RoboDK station: kuka_frame.rdk

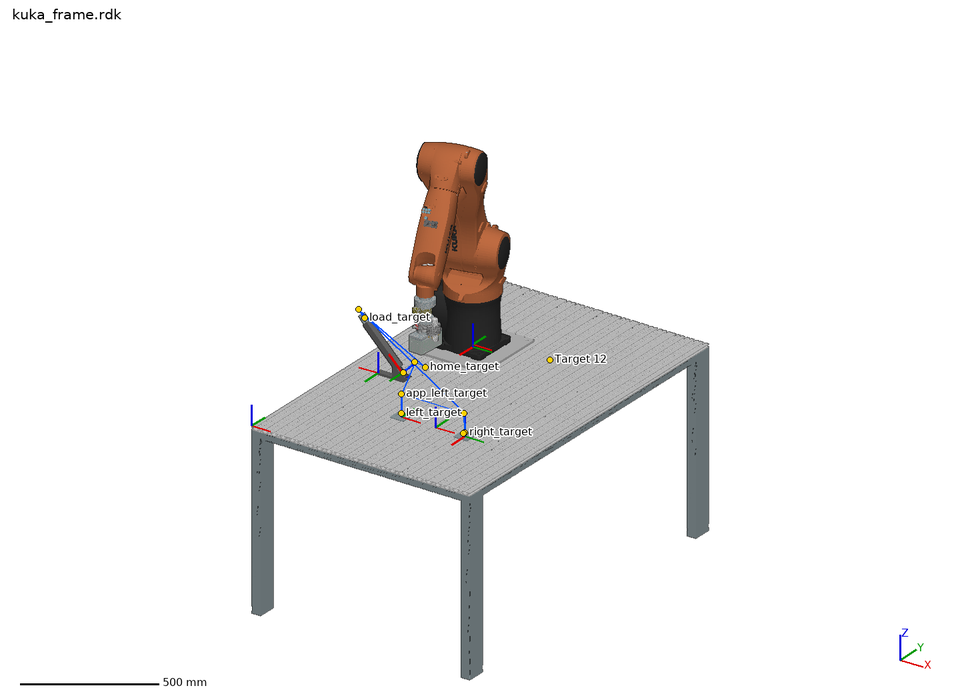
[picture v0: the station drawn from its stored meshes, robots at their saved joint values, targets as dots, program paths as lines]
Station kuka_frame(vansh2) (saved by RoboDK 5.8.0). Poses are relative to the parent item; angles as X-Y-Z fixed-axis rotations.
Station parameters (name, value as stored): LIN64
  - frame table_frame at (0, 0, 0) mm
    - object table_object at (0, 0, 0) mm, size 960.1 x 1500 x 750 mm, geometry from table_object.sld
    - frame base_plate_frame at (280, 990, 0) mm, rotated rx 0 ry 0 rz -90 deg
      - object base_plate_object at (0, 0, 0) mm, size 320 x 320 x 10 mm, geometry from base_plate_object.sld
    - frame slider_frame at (125, 617, 0) mm, rotated rx 0 ry 0 rz 180 deg
      - object slider_object at (0, 0, 0) mm, size 198.7 x 26 x 198.7 mm, 1 curves, geometry from slider_object.sld
    - frame slider_parts_frame at (232.7, 617, 30.7) mm, rotated rx 0 ry -45 rz 180 deg
    - frame pickanddrop at (550, 370, 0) mm
    - frame right_frame at (680, 370, 0) mm, rotated rx 0 ry 0 rz -90 deg
      - object right_plate_object at (0, 0, 0) mm, size 60 x 60 x 9 mm, 1 curves, geometry from right_plate_object.sld
    - frame left_frame at (400, 370, 0) mm
      - object left_plate_object at (0, 0, 0) mm, size 60 x 60 x 9 mm, 1 curves, geometry from left_plate_object.sld
    - frame kuka_frame at (280, 990, 10) mm
      - robot KUKA KR 6 R900 sixx: 6 axes, payload 6 kg, reach 901 mm, repeatability 0.03 mm, weight 52 kg
          modified DH rows (alpha deg, a mm, theta deg, d mm): 0, 0, 0, 400; -90, 25, 0, 0; 0, 455, -90, 0; -90, 35, 0, 420; 90, 0, 0, 0; -90, 0, 180, 80
          joint limits [-170, -190, -120, -185, -120, -350] to [170, 45, 156, 185, 120, 350]; home [0, -90, 90, 0, 0, 0]; saved at [75.683, -66.176, 119.978, 0, 36.199, -61.317]
        - robot gripper: 1 axes
            joint limits [0] to [50]; home [0]; saved at [50]
        - tool gripper_tcp, TCP at (0, 0, 288) mm, rotated rx 0 ry 0 rz 43 deg
    - target home_target (Cartesian target) at (399.96, 519.99, 139.97) mm, rotated rx -180 ry 0 rz 0 deg; joints [75.683, -66.176, 119.978, 0, 36.199, -61.317] of KUKA KR 6 R900 sixx
    - target left_target (Cartesian target) at (400, 370, 15) mm, rotated rx -180 ry 0 rz 0 deg; joints [79.046, -41.366, 97.165, 0, 34.201, -57.954] of KUKA KR 6 R900 sixx
    - target app_left_target (Cartesian target) at (400, 370, 93) mm, rotated rx -180 ry 0 rz 0 deg; joints [79.046, -48.593, 96.885, 0, 41.708, -57.954] of KUKA KR 6 R900 sixx
    - target right_target (Cartesian target) at (680, 370, 15) mm, rotated rx -180 ry 0 rz -90 deg; joints [57.171, -31.816, 75.866, 0, 45.949, -169.829] of KUKA KR 6 R900 sixx
    - target app_right_target (Cartesian target) at (676.53, 370, 93) mm, rotated rx -180 ry 0 rz -180 deg; joints [57.398, -38.147, 75.992, 0, 52.155, 100.398] of KUKA KR 6 R900 sixx
    - target slider_part_target (Cartesian target) at (234.82, 617, 32.82) mm, rotated rx 180 ry 45 rz 0 deg; joints [60.036, -41.203, 127.341, 56.857, 47.023, -132.424] of KUKA KR 6 R900 sixx
    - target app_sliderpart_target (Cartesian target) at (286, 617, 88.78) mm, rotated rx -180 ry 50 rz 0 deg; joints [52.337, -44.49, 122.484, 45.711, 57.903, -125.791] of KUKA KR 6 R900 sixx
    - target load_target (Cartesian target) at (66.24, 617, 203.91) mm, rotated rx -180 ry 50 rz 0 deg; joints [79.647, -66.13, 137.097, 65.731, 55.754, -114.165] of KUKA KR 6 R900 sixx
    - target app_load_target (Cartesian target) at (38.79, 617, 231.21) mm, rotated rx 180 ry 49 rz 0 deg; joints [84.408, -71.376, 137.116, 65.861, 55.395, -107.211] of KUKA KR 6 R900 sixx
    - target open_grip (joint target) at (399.96, 519.99, -148.03) mm, rotated rx -180 ry 0 rz -43 deg; joints [50] of gripper
    - target close_grippertarget (joint target) at (399.96, 519.99, -148.03) mm, rotated rx -180 ry 0 rz -43 deg; joints [20, -66.176, 119.978, -180, -36.199, 118.683] of gripper
    - target Target 12 (Cartesian target) at (735.82, 824.09, 139.97) mm, rotated rx -180 ry 0 rz 55.68 deg; joints [20, -66.176, 119.978, 0, 36.199, 298.683] of KUKA KR 6 R900 sixx
    - target Target 13 (Cartesian target) at (735.82, 824.09, 139.97) mm, rotated rx -180 ry 0 rz 55.68 deg; joints [20, -66.176, 119.978, 0, 36.199, 298.683] of KUKA KR 6 R900 sixx
    - target Target 14 (Cartesian target) at (735.82, 824.09, 139.97) mm, rotated rx -180 ry 0 rz 55.68 deg; joints [20, -66.176, 119.978, 0, 36.199, 298.683] of KUKA KR 6 R900 sixx
    - target Target 15 (Cartesian target) at (735.82, 824.09, 139.97) mm, rotated rx -180 ry 0 rz 55.68 deg; joints [20, -66.176, 119.978, 0, 36.199, 298.683] of KUKA KR 6 R900 sixx
    - target Target 16 (Cartesian target) at (735.82, 824.09, 139.97) mm, rotated rx -180 ry 0 rz 55.68 deg; joints [20, -66.176, 119.978, 0, 36.199, 298.683] of KUKA KR 6 R900 sixx
    - target Target 17 (Cartesian target) at (735.82, 824.09, 139.97) mm, rotated rx -180 ry 0 rz 55.68 deg; joints [20, -66.176, 119.978, 0, 36.199, 298.683] of KUKA KR 6 R900 sixx
    - target Target 18 (Cartesian target) at (735.82, 824.09, 139.97) mm, rotated rx -180 ry 0 rz 55.68 deg; joints [20, -66.176, 119.978, 0, 36.199, 298.683] of KUKA KR 6 R900 sixx
    - target Target 19 (Cartesian target) at (735.82, 824.09, 139.97) mm, rotated rx -180 ry 0 rz 55.68 deg; joints [20, -66.176, 119.978, 0, 36.199, 298.683] of KUKA KR 6 R900 sixx
    - target Target 20 (Cartesian target) at (735.82, 824.09, 139.97) mm, rotated rx -180 ry 0 rz 55.68 deg; joints [20, -66.176, 119.978, 0, 36.199, 298.683] of KUKA KR 6 R900 sixx
    - target Target 21 (Cartesian target) at (735.82, 824.09, 139.97) mm, rotated rx -180 ry 0 rz 55.68 deg; joints [20, -66.176, 119.978, 0, 36.199, 298.683] of KUKA KR 6 R900 sixx
    - target Target 22 (Cartesian target) at (735.82, 824.09, 139.97) mm, rotated rx -180 ry 0 rz 55.68 deg; joints [20, -66.176, 119.978, 0, 36.199, 298.683] of KUKA KR 6 R900 sixx
    - target Target 23 (Cartesian target) at (735.82, 824.09, 139.97) mm, rotated rx -180 ry 0 rz 55.68 deg; joints [20, -66.176, 119.978, 0, 36.199, 298.683] of KUKA KR 6 R900 sixx
    - target Target 24 (Cartesian target) at (735.82, 824.09, 139.97) mm, rotated rx -180 ry 0 rz 55.68 deg; joints [20, -66.176, 119.978, 0, 36.199, 298.683] of KUKA KR 6 R900 sixx
    - target Target 25 (Cartesian target) at (735.82, 824.09, 139.97) mm, rotated rx -180 ry 0 rz 55.68 deg; joints [20, -66.176, 119.978, 0, 36.199, 298.683] of KUKA KR 6 R900 sixx
    - target Target 26 (Cartesian target) at (735.82, 824.09, 139.97) mm, rotated rx -180 ry 0 rz 55.68 deg; joints [20, -66.176, 119.978, 0, 36.199, 298.683] of KUKA KR 6 R900 sixx
    - target Target 27 (Cartesian target) at (735.82, 824.09, 139.97) mm, rotated rx -180 ry 0 rz 55.68 deg; joints [20, -66.176, 119.978, 0, 36.199, 298.683] of KUKA KR 6 R900 sixx
    - target Target 28 (Cartesian target) at (735.82, 824.09, 139.97) mm, rotated rx -180 ry 0 rz 55.68 deg; joints [20, -66.176, 119.978, 0, 36.199, 298.683] of KUKA KR 6 R900 sixx
    - target Target 29 (Cartesian target) at (735.82, 824.09, 139.97) mm, rotated rx -180 ry 0 rz 55.68 deg; joints [20, -66.176, 119.978, 0, 36.199, 298.683] of KUKA KR 6 R900 sixx
    - target Target 30 (Cartesian target) at (676.53, 364.14, 15) mm, rotated rx -180 ry 0 rz -90 deg; joints [57.643, -31.498, 75.173, 0, 46.325, -169.357] of KUKA KR 6 R900 sixx
    - target Target 31 (Cartesian target) at (676.53, 364.14, 15) mm, rotated rx -180 ry 0 rz -90 deg; joints [57.643, -31.498, 75.173, 0, 46.325, -169.357] of KUKA KR 6 R900 sixx
  - folder programs
    - program factory_reset (1 instructions, listed below)
    - program open_gripper (1 instructions, listed below)
    - program close_gripper (2 instructions, listed below)
    - program main (34 instructions, listed below)
  - object part_object at (63.46, 617, 201.02) mm, rotated rx 0 ry -50 rz -180 deg, size 40 x 20 x 20 mm, 1 curves, geometry from part_object.sld
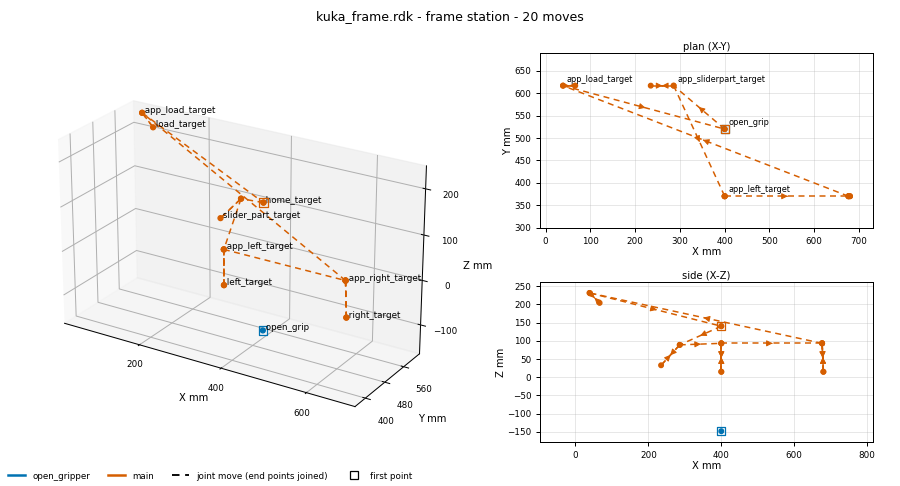
[picture p0: tool path of kuka_frame.rdk in frame station, 20 of 20 moves have a stored position in this frame; points joined in program order, loops and branches not executed]

--- program factory_reset (robot KUKA KR 6 R900 sixx) ---
  Replace objects

--- program open_gripper (robot gripper) ---
  MoveJ (open_grip)

--- program close_gripper (robot gripper) ---
  Set Ref.: table_frame
  Set Tool: gripper_tcp

--- program main (robot KUKA KR 6 R900 sixx) ---
  Set Ref.: table_frame
  Set Tool: gripper_tcp
  Call open_gripper
  MoveJ (home_target)
  MoveJ (app_sliderpart_target)
  MoveJ (slider_part_target)
  Call close_gripper
  Attach to gripper_tcp
  MoveJ (app_sliderpart_target)
  MoveJ (app_left_target)
  MoveJ (left_target)
  Call open_gripper
  Detach from gripper_tcp
  MoveJ (app_left_target)
  MoveJ (left_target)
  Call close_gripper
  Attach to gripper_tcp
  MoveJ (app_left_target)
  MoveJ (app_right_target)
  MoveJ (right_target)
  Call open_gripper
  Detach from gripper_tcp
  MoveJ (app_right_target)
  MoveJ (right_target)
  Call close_gripper
  Attach to gripper_tcp
  MoveJ (app_right_target)
  MoveJ (app_right_target)
  MoveJ (app_load_target)
  MoveJ (load_target)
  Call open_gripper
  Detach from gripper_tcp
  MoveJ (app_load_target)
  MoveJ (home_target)
